  MoveL 647 to (-2817.75, 812.38, 1030.88) mm, rotated rx -103.17 ry -2.27 rz -179.99 deg; joints [-49.243, 2.601, 19.186, -115.031, 26.585, 9.042, -170]
  MoveL 648 to (-2817.75, 831.47, 992.27) mm, rotated rx -103.22 ry -3.45 rz -179.99 deg; joints [-48.787, 2.468, 20.52, -112.558, 24.893, 6.606, -170]
  MoveL 649 to (-2817.75, 844.77, 965.38) mm, rotated rx -103.26 ry -4.26 rz -179.99 deg; joints [-48.461, 2.4, 21.424, -110.645, 23.624, 4.8, -170]
  MoveL 650 to (-2817.75, 844.7, 935.74) mm, rotated rx -99.91 ry -3.73 rz -179.99 deg; joints [-48.443, 3.334, 22.932, -110.863, 27.836, -0.78, -170]
  MoveL 651 to (-2817.75, 844.62, 905.74) mm, rotated rx -96.49 ry -2.63 rz -179.99 deg; joints [-48.478, 4.555, 24.383, -112.634, 33.789, -5.769, -170]
  MoveL 652 to (-2817.75, 844.55, 875.74) mm, rotated rx -93.08 ry 1.03 rz 180 deg; joints [-48.572, 6.332, 25.892, -116.809, 44.188, -9.974, -170]
  MoveL 653 to (-2817.75, 844.47, 845.74) mm, rotated rx -89.7 ry 0.4 rz -179.6 deg; joints [-48.723, 7.85, 26.739, -119.615, 48.753, -14.494, -170]
  MoveL 654 to (-2817.75, 844.3, 816.11) mm, rotated rx -89.68 ry 0.41 rz -179.59 deg; joints [-48.729, 8.688, 27.11, -120.262, 50.179, -15.333, -170]
  MoveL 655 to (-2817.75, 844.12, 786.11) mm, rotated rx -89.67 ry 0.42 rz -179.58 deg; joints [-48.736, 9.565, 27.459, -120.936, 51.634, -16.183, -170]
  MoveL 656 to (-2817.75, 843.95, 756.11) mm, rotated rx -89.65 ry 0.43 rz -179.57 deg; joints [-48.743, 10.47, 27.78, -121.627, 53.1, -17.032, -170]
  MoveL 657 to (-2817.75, 843.77, 726.11) mm, rotated rx -89.64 ry 0.45 rz -179.56 deg; joints [-48.751, 11.401, 28.074, -122.336, 54.575, -17.882, -170]
  MoveL 658 to (-2817.75, 843.58, 696.48) mm, rotated rx -89.64 ry 0.45 rz -179.55 deg; joints [-48.758, 12.343, 28.335, -123.033, 56.012, -18.708, -170]
  MoveL 659 to (-2817.75, 843.38, 666.48) mm, rotated rx -89.64 ry 0.46 rz -179.54 deg; joints [-48.765, 13.323, 28.571, -123.754, 57.474, -19.544, -170]
  MoveL 660 to (-2817.75, 843.19, 636.48) mm, rotated rx -89.64 ry 0.47 rz -179.53 deg; joints [-48.773, 14.327, 28.78, -124.49, 58.942, -20.381, -170]
  MoveL 661 to (-2817.75, 843, 606.48) mm, rotated rx -89.64 ry 0.48 rz -179.52 deg; joints [-48.782, 15.356, 28.96, -125.239, 60.414, -21.219, -170]
  MoveL 662 to (-2817.75, 842.82, 569.69) mm, rotated rx -89.65 ry 0.48 rz -179.52 deg; joints [-48.789, 16.643, 29.145, -126.15, 62.194, -22.238, -170]
  MoveL 663 to (-2817.75, 842.68, 539.69) mm, rotated rx -89.66 ry 0.49 rz -179.51 deg; joints [-48.796, 17.718, 29.264, -126.907, 63.648, -23.068, -170]
  MoveL 664 to (-2817.75, 842.54, 509.69) mm, rotated rx -89.67 ry 0.49 rz -179.51 deg; joints [-48.803, 18.815, 29.354, -127.675, 65.102, -23.898, -170]
  MoveL 665 to (-2817.75, 842.4, 479.69) mm, rotated rx -89.68 ry 0.5 rz -179.5 deg; joints [-48.811, 19.933, 29.417, -128.453, 66.555, -24.728, -170]
  MoveL 666 to (-2817.75, 842.26, 449.69) mm, rotated rx -89.69 ry 0.5 rz -179.5 deg; joints [-48.819, 21.072, 29.451, -129.241, 68.007, -25.558, -170]
  MoveL 667 to (-2817.75, 842.12, 419.69) mm, rotated rx -89.7 ry 0.51 rz -179.5 deg; joints [-48.827, 22.229, 29.456, -130.038, 69.455, -26.387, -170]
  MoveL 668 to (-2817.75, 841.97, 389.69) mm, rotated rx -89.71 ry 0.51 rz -179.49 deg; joints [-48.836, 23.406, 29.433, -130.843, 70.899, -27.214, -170]
  MoveL 669 to (-2817.75, 841.83, 359.69) mm, rotated rx -89.73 ry 0.52 rz -179.49 deg; joints [-48.845, 24.599, 29.381, -131.655, 72.337, -28.04, -170]
  MoveL 670 to (-2817.75, 841.69, 329.69) mm, rotated rx -89.74 ry 0.52 rz -179.48 deg; joints [-48.855, 25.809, 29.301, -132.473, 73.767, -28.864, -170]
  MoveL 671 to (-2817.75, 841.54, 299.69) mm, rotated rx -89.75 ry 0.52 rz -179.48 deg; joints [-48.865, 27.035, 29.193, -133.296, 75.189, -29.685, -170]
  MoveL 672 to (-2817.75, 841.4, 269.7) mm, rotated rx -89.76 ry 0.53 rz -179.47 deg; joints [-48.876, 28.275, 29.056, -134.124, 76.601, -30.503, -170]
  MoveL 673 to (-2817.75, 841.26, 239.69) mm, rotated rx -89.75 ry -19.47 rz -179.55 deg; joints [-47.931, 25.571, 28.432, -109.218, 40.774, -38.612, -170]
  MoveL 674 to (-2817.75, 841.12, 209.69) mm, rotated rx -89.77 ry -19.46 rz -179.54 deg; joints [-47.933, 26.785, 28.338, -110.005, 42.222, -39.195, -170]
  MoveL 675 to (-2817.75, 841.08, 201.69) mm, rotated rx -89.77 ry -19.46 rz -179.54 deg; joints [-47.932, 27.113, 28.308, -110.208, 42.604, -39.356, -170]
  Set speed (1000.0 mm/s)
  MoveL 676 to (-2817.75, 841.08, 201.69) mm, rotated rx -89.77 ry -19.46 rz -179.54 deg; joints [-47.932, 27.113, 28.308, -110.208, 42.604, -39.356, -170]
  MoveL 677 to (-2818.68, 941.08, 201.3) mm, rotated rx -89.77 ry -19.46 rz -179.54 deg; joints [-46.038, 24.56, 32.438, -107.449, 43.1, -41.713, -170]
  Set speed (1000.0 mm/s)
  MoveL 678 to (-2898.69, 940.29, 202.16) mm, rotated rx -89.77 ry -19.46 rz -179.54 deg; joints [-49.032, 23.561, 34.225, -114.018, 46.527, -39.844, -170]
  MoveL 679 to (-2897.75, 840.3, 202.54) mm, rotated rx -89.77 ry -19.46 rz -179.54 deg; joints [-50.794, 26.176, 30.018, -116.607, 46.068, -37.565, -170]
  MoveL 680 to (-2897.75, 840.3, 202.54) mm, rotated rx -89.77 ry -19.46 rz -179.54 deg; joints [-50.794, 26.176, 30.018, -116.607, 46.068, -37.565, -170]
  Set speed (50.0 mm/s)
  MoveL 681 to (-2897.75, 840.33, 210.54) mm, rotated rx -89.77 ry -19.46 rz -179.54 deg; joints [-50.794, 25.842, 30.05, -116.45, 45.715, -37.364, -170]
  MoveL 682 to (-2897.75, 840.45, 240.54) mm, rotated rx -89.75 ry -19.46 rz -179.55 deg; joints [-50.792, 24.603, 30.15, -115.833, 44.378, -36.641, -170]
  MoveL 683 to (-2897.75, 840.57, 270.54) mm, rotated rx -89.74 ry -19.47 rz -179.56 deg; joints [-50.792, 23.378, 30.221, -115.24, 43.04, -35.89, -170]
  MoveL 684 to (-2897.75, 840.7, 300.54) mm, rotated rx -89.73 ry -19.47 rz -179.56 deg; joints [-50.792, 22.17, 30.264, -114.657, 41.697, -35.129, -170]
  MoveL 685 to (-2897.75, 840.81, 330.55) mm, rotated rx -89.74 ry 0.53 rz -179.48 deg; joints [-51.786, 24.874, 30.905, -137.578, 76.653, -28.084, -170]
  MoveL 686 to (-2897.75, 840.94, 360.54) mm, rotated rx -89.73 ry 0.52 rz -179.48 deg; joints [-51.777, 23.638, 30.987, -136.808, 75.263, -27.171, -170]
  MoveL 687 to (-2897.75, 841.02, 380.87) mm, rotated rx -89.72 ry 0.52 rz -179.48 deg; joints [-51.771, 22.81, 31.027, -136.292, 74.318, -26.55, -170]
  MoveL 688 to (-2897.75, 841.2, 410.87) mm, rotated rx -89.71 ry 0.52 rz -179.49 deg; joints [-51.761, 21.603, 31.063, -135.536, 72.922, -25.638, -170]
  MoveL 689 to (-2897.75, 841.38, 440.87) mm, rotated rx -89.7 ry 0.51 rz -179.49 deg; joints [-51.751, 20.414, 31.07, -134.791, 71.523, -24.724, -170]
  MoveL 690 to (-2897.75, 841.55, 470.87) mm, rotated rx -89.68 ry 0.51 rz -179.5 deg; joints [-51.742, 19.245, 31.049, -134.059, 70.124, -23.807, -170]
  MoveL 691 to (-2897.75, 841.73, 500.87) mm, rotated rx -89.67 ry 0.5 rz -179.5 deg; joints [-51.734, 18.096, 30.999, -133.341, 68.725, -22.888, -170]
  MoveL 692 to (-2897.75, 841.9, 530.87) mm, rotated rx -89.65 ry 0.5 rz -179.51 deg; joints [-51.726, 16.969, 30.92, -132.638, 67.328, -21.966, -170]
  MoveL 693 to (-2897.75, 842.07, 560.87) mm, rotated rx -89.64 ry 0.49 rz -179.51 deg; joints [-51.718, 15.864, 30.813, -131.95, 65.935, -21.042, -170]
  MoveL 694 to (-2897.75, 842.25, 590.87) mm, rotated rx -89.63 ry 0.48 rz -179.52 deg; joints [-51.711, 14.782, 30.677, -131.28, 64.547, -20.117, -170]
  MoveL 695 to (-2897.75, 842.37, 611.21) mm, rotated rx -89.62 ry 0.48 rz -179.52 deg; joints [-51.707, 14.062, 30.568, -130.835, 63.609, -19.488, -170]
  MoveL 696 to (-2897.75, 842.57, 641.21) mm, rotated rx -89.62 ry 0.47 rz -179.53 deg; joints [-51.699, 13.016, 30.385, -130.177, 62.209, -18.547, -170]
  MoveL 697 to (-2897.75, 842.78, 671.2) mm, rotated rx -89.62 ry 0.46 rz -179.54 deg; joints [-51.692, 11.994, 30.174, -129.54, 60.818, -17.604, -170]
  MoveL 698 to (-2897.75, 842.98, 701.2) mm, rotated rx -89.61 ry 0.46 rz -179.55 deg; joints [-51.685, 10.999, 29.935, -128.923, 59.438, -16.66, -170]
  MoveL 699 to (-2897.75, 843.19, 731.86) mm, rotated rx -89.61 ry 0.45 rz -179.55 deg; joints [-51.678, 10.01, 29.661, -128.315, 58.039, -15.693, -170]
  MoveL 700 to (-2897.75, 843.38, 761.86) mm, rotated rx -89.63 ry 0.44 rz -179.57 deg; joints [-51.671, 9.065, 29.363, -127.726, 56.658, -14.729, -170]
  MoveL 701 to (-2897.75, 843.57, 791.85) mm, rotated rx -89.64 ry 0.43 rz -179.58 deg; joints [-51.665, 8.149, 29.038, -127.162, 55.292, -13.763, -170]
  MoveL 702 to (-2897.75, 843.76, 821.85) mm, rotated rx -89.65 ry 0.41 rz -179.59 deg; joints [-51.659, 7.261, 28.685, -126.623, 53.941, -12.795, -170]
  MoveL 703 to (-2897.75, 843.96, 852.51) mm, rotated rx -89.67 ry 0.4 rz -179.6 deg; joints [-51.653, 6.383, 28.296, -126.1, 52.579, -11.802, -170]
  MoveL 704 to (-2897.75, 844.05, 882.51) mm, rotated rx -93.14 ry 0.91 rz 180 deg; joints [-51.496, 4.806, 27.427, -123.67, 48.036, -6.803, -170]
  MoveL 705 to (-2897.75, 844.14, 912.51) mm, rotated rx -96.65 ry -2.69 rz -179.99 deg; joints [-51.402, 3.012, 25.922, -121.089, 38.685, -1.519, -170]
  MoveL 706 to (-2897.75, 844.24, 942.51) mm, rotated rx -100.16 ry -3.78 rz -179.99 deg; joints [-51.372, 1.784, 24.461, -120.72, 33.653, 4.42, -170]
  MoveL 707 to (-2897.75, 844.33, 973.16) mm, rotated rx -103.72 ry -4.31 rz -179.99 deg; joints [-51.402, 0.829, 22.882, -121.934, 30.285, 11.118, -170]
  MoveL 708 to (-2897.75, 830.58, 999.82) mm, rotated rx -103.69 ry -3.5 rz -179.99 deg; joints [-51.725, 0.942, 21.926, -123.457, 31.388, 12.672, -170]
  MoveL 709 to (-2897.75, 809.97, 1039.78) mm, rotated rx -103.64 ry -2.29 rz -179.99 deg; joints [-52.194, 1.149, 20.461, -125.527, 32.941, 14.887, -170]
  MoveL 710 to (-2897.75, 796.37, 1066.52) mm, rotated rx -108.84 ry -1.41 rz -180 deg; joints [-52.753, 1.175, 17.955, -130.919, 33.223, 25.392, -170]
  MoveL 711 to (-2897.75, 775.99, 1106.6) mm, rotated rx -116.66 ry -0.72 rz -180 deg; joints [-53.755, 1.801, 13.687, -142.342, 36.014, 42.395, -170]
  MoveL 712 to (-2897.75, 762.7, 1133.49) mm, rotated rx -116.26 ry 0.34 rz 180 deg; joints [-54.078, 2.014, 12.796, -142.876, 37.16, 42.843, -170]
  MoveL 713 to (-2897.75, 749.89, 1159.4) mm, rotated rx -115.89 ry 1.39 rz 180 deg; joints [-54.38, 2.235, 11.926, -143.28, 38.216, 43.237, -170]
  MoveL 714 to (-2897.75, 746.94, 1165.63) mm, rotated rx -115.75 ry 1.69 rz 180 deg; joints [-54.45, 2.282, 11.747, -143.268, 38.475, 43.216, -170]
  Set speed (1000.0 mm/s)
  MoveL 715 to (-2897.75, 746.94, 1165.63) mm, rotated rx -115.75 ry 1.69 rz 180 deg; joints [-54.45, 2.282, 11.747, -143.268, 38.475, 43.216, -170]
  MoveL 716 to (-2899.02, 837.01, 1209.06) mm, rotated rx -115.75 ry 1.69 rz 180 deg; joints [-53.221, -1.859, 14.256, -141.506, 35.807, 44.207, -170]
  Set speed (1000.0 mm/s)
  MoveL 717 to (-2979.82, 828.97, 1222.94) mm, rotated rx -116.54 ry 2.68 rz 179.99 deg; joints [-56.639, -2.784, 14.766, -150.413, 43.399, 48.713, -170]
  MoveL 718 to (-2977.75, 739.51, 1178.3) mm, rotated rx -116.54 ry 2.68 rz 179.99 deg; joints [-57.642, 1.416, 12.276, -151.236, 45.388, 47.167, -170]
  MoveL 719 to (-2977.75, 739.51, 1178.3) mm, rotated rx -116.54 ry 2.68 rz 179.99 deg; joints [-57.642, 1.416, 12.276, -151.236, 45.388, 47.167, -170]
  Set speed (50.0 mm/s)
  MoveL 720 to (-2977.75, 743.33, 1170.64) mm, rotated rx -116.9 ry 1.76 rz 180 deg; joints [-57.513, 1.36, 12.335, -151.884, 44.805, 47.788, -170]
  MoveL 721 to (-2977.75, 757.4, 1143.51) mm, rotated rx -117.39 ry 0.32 rz 180 deg; joints [-57.172, 1.086, 13.2, -151.998, 43.61, 47.787, -170]
  MoveL 722 to (-2977.75, 771.22, 1116.88) mm, rotated rx -117.73 ry -0.71 rz -180 deg; joints [-56.858, 0.82, 14.158, -151.612, 42.569, 47.354, -170]
  MoveL 723 to (-2977.75, 779.23, 1101.8) mm, rotated rx -114.73 ry -0.91 rz -180 deg; joints [-56.469, 0.423, 15.935, -147.19, 41.112, 41.102, -170]
  MoveL 724 to (-2977.75, 793.31, 1075.31) mm, rotated rx -109.41 ry -1.43 rz -180 deg; joints [-55.836, -0.019, 18.855, -140.279, 39.466, 30.188, -170]
  MoveL 725 to (-2977.75, 807.39, 1048.82) mm, rotated rx -104.13 ry -2.31 rz -179.99 deg; joints [-55.283, -0.138, 21.477, -134.908, 38.92, 19.784, -170]
  MoveL 726 to (-2977.75, 815.48, 1033.78) mm, rotated rx -104.14 ry -2.76 rz -179.99 deg; joints [-55.114, -0.249, 22.065, -134.286, 38.393, 19.044, -170]
  MoveL 727 to (-2977.75, 829.69, 1007.36) mm, rotated rx -104.17 ry -3.56 rz -179.99 deg; joints [-54.811, -0.429, 23.083, -133.124, 37.432, 17.709, -170]
  MoveL 728 to (-2977.75, 843.89, 980.94) mm, rotated rx -104.2 ry -4.35 rz -179.99 deg; joints [-54.498, -0.589, 24.085, -131.869, 36.428, 16.329, -170]
  MoveL 729 to (-2977.75, 843.78, 949.27) mm, rotated rx -100.41 ry -3.82 rz -179.99 deg; joints [-54.457, 0.383, 25.761, -129.756, 39.228, 8.855, -170]
  MoveL 730 to (-2977.75, 843.66, 919.27) mm, rotated rx -96.8 ry -2.76 rz -179.99 deg; joints [-54.481, 1.615, 27.246, -129.178, 43.575, 2.269, -170]
  MoveL 731 to (-2977.75, 843.55, 889.27) mm, rotated rx -93.2 ry 0.78 rz 180 deg; joints [-54.569, 3.423, 28.761, -130.525, 52.047, -3.846, -170]
  MoveL 732 to (-2977.75, 843.44, 859.27) mm, rotated rx -89.64 ry 0.41 rz -179.6 deg; joints [-54.731, 5.056, 29.653, -132.597, 56.549, -9.299, -170]
  MoveL 733 to (-2977.75, 843.22, 827.6) mm, rotated rx -89.62 ry 0.42 rz -179.58 deg; joints [-54.735, 5.97, 30.06, -133.01, 57.842, -10.434, -170]
  MoveL 734 to (-2977.75, 843.02, 797.6) mm, rotated rx -89.61 ry 0.43 rz -179.57 deg; joints [-54.739, 6.868, 30.418, -133.433, 59.089, -11.505, -170]
  MoveL 735 to (-2977.75, 842.81, 767.6) mm, rotated rx -89.6 ry 0.44 rz -179.56 deg; joints [-54.744, 7.794, 30.748, -133.887, 60.356, -12.572, -170]
  MoveL 736 to (-2977.75, 842.61, 737.6) mm, rotated rx -89.59 ry 0.45 rz -179.55 deg; joints [-54.75, 8.75, 31.05, -134.37, 61.641, -13.636, -170]
  MoveL 737 to (-2977.75, 842.38, 705.93) mm, rotated rx -89.59 ry 0.46 rz -179.54 deg; joints [-54.756, 9.785, 31.337, -134.893, 62.992, -14.739, -170]
  MoveL 738 to (-2977.75, 842.16, 675.93) mm, rotated rx -89.59 ry 0.47 rz -179.53 deg; joints [-54.761, 10.794, 31.58, -135.416, 64.287, -15.781, -170]
  MoveL 739 to (-2977.75, 841.95, 645.94) mm, rotated rx -89.6 ry 0.48 rz -179.53 deg; joints [-54.768, 11.83, 31.795, -135.965, 65.597, -16.82, -170]
  MoveL 740 to (-2977.75, 841.73, 615.94) mm, rotated rx -89.6 ry 0.48 rz -179.52 deg; joints [-54.775, 12.893, 31.981, -136.537, 66.918, -17.856, -170]
  MoveL 741 to (-2977.75, 841.6, 593.66) mm, rotated rx -89.61 ry 0.49 rz -179.51 deg; joints [-54.779, 13.694, 32.101, -136.965, 67.89, -18.613, -170]
  MoveL 742 to (-2977.75, 841.41, 563.66) mm, rotated rx -89.62 ry 0.49 rz -179.51 deg; joints [-54.786, 14.794, 32.238, -137.56, 69.208, -19.63, -170]
  MoveL 743 to (-2977.75, 841.23, 533.66) mm, rotated rx -89.64 ry 0.5 rz -179.51 deg; joints [-54.792, 15.918, 32.346, -138.176, 70.533, -20.644, -170]
  MoveL 744 to (-2977.75, 841.05, 503.66) mm, rotated rx -89.65 ry 0.5 rz -179.5 deg; joints [-54.8, 17.065, 32.425, -138.812, 71.866, -21.655, -170]
  MoveL 745 to (-2977.75, 840.87, 473.66) mm, rotated rx -89.67 ry 0.51 rz -179.5 deg; joints [-54.808, 18.234, 32.475, -139.466, 73.203, -22.662, -170]
  MoveL 746 to (-2977.75, 840.68, 443.66) mm, rotated rx -89.68 ry 0.51 rz -179.49 deg; joints [-54.817, 19.425, 32.496, -140.138, 74.543, -23.665, -170]
  MoveL 747 to (-2977.75, 840.49, 413.67) mm, rotated rx -89.7 ry 0.52 rz -179.49 deg; joints [-54.826, 20.635, 32.488, -140.826, 75.886, -24.664, -170]
  MoveL 748 to (-2977.75, 840.31, 383.68) mm, rotated rx -89.71 ry 0.52 rz -179.48 deg; joints [-54.836, 21.864, 32.45, -141.528, 77.228, -25.659, -170]
  MoveL 749 to (-2977.75, 840.22, 361.39) mm, rotated rx -89.7 ry -19.48 rz -179.58 deg; joints [-53.805, 18.856, 31.81, -120.744, 43.029, -31.253, -170]
  MoveL 750 to (-2977.75, 840.1, 331.39) mm, rotated rx -89.71 ry -19.47 rz -179.57 deg; joints [-53.802, 20.05, 31.819, -121.094, 44.23, -32.192, -170]
  MoveL 751 to (-2977.75, 839.97, 301.39) mm, rotated rx -89.72 ry -19.47 rz -179.57 deg; joints [-53.8, 21.263, 31.798, -121.472, 45.44, -33.114, -170]
  MoveL 752 to (-2977.75, 839.84, 271.39) mm, rotated rx -89.73 ry -19.47 rz -179.56 deg; joints [-53.798, 22.495, 31.75, -121.875, 46.657, -34.019, -170]
  MoveL 753 to (-2977.75, 839.71, 241.39) mm, rotated rx -89.74 ry -19.46 rz -179.55 deg; joints [-53.797, 23.744, 31.672, -122.3, 47.878, -34.907, -170]
  MoveL 754 to (-2977.75, 839.58, 211.39) mm, rotated rx -89.75 ry -19.46 rz -179.55 deg; joints [-53.796, 25.01, 31.566, -122.744, 49.101, -35.779, -170]
  MoveL 755 to (-2977.75, 839.55, 203.39) mm, rotated rx -89.75 ry -19.46 rz -179.55 deg; joints [-53.795, 25.351, 31.533, -122.862, 49.427, -36.014, -170]
  Set speed (1000.0 mm/s)
  MoveL 756 to (-2977.75, 839.55, 203.39) mm, rotated rx -89.75 ry -19.46 rz -179.55 deg; joints [-53.795, 25.351, 31.533, -122.862, 49.427, -36.014, -170]
  MoveL 757 to (-2978.68, 939.54, 202.98) mm, rotated rx -89.75 ry -19.46 rz -179.55 deg; joints [-52.193, 22.678, 35.815, -120.489, 49.872, -38.211, -170]
  Set speed (1000.0 mm/s)
  MoveL 758 to (-3058.69, 938.8, 203.83) mm, rotated rx -89.75 ry -19.46 rz -179.54 deg; joints [-55.525, 21.905, 37.195, -126.964, 53.169, -36.713, -170]
  MoveL 759 to (-3057.75, 838.8, 204.24) mm, rotated rx -89.75 ry -19.46 rz -179.54 deg; joints [-56.937, 24.633, 32.844, -129.079, 52.722, -34.6, -170]
  MoveL 760 to (-3057.75, 838.8, 204.24) mm, rotated rx -89.75 ry -19.46 rz -179.54 deg; joints [-56.937, 24.633, 32.844, -129.079, 52.722, -34.6, -170]
  Set speed (50.0 mm/s)
  MoveL 761 to (-3057.75, 838.84, 212.24) mm, rotated rx -89.75 ry -19.46 rz -179.54 deg; joints [-56.939, 24.287, 32.878, -128.997, 52.425, -34.335, -170]
  MoveL 762 to (-3057.75, 838.97, 242.24) mm, rotated rx -89.73 ry -19.46 rz -179.56 deg; joints [-56.94, 23.001, 32.989, -128.679, 51.31, -33.367, -170]
  MoveL 763 to (-3057.75, 839.11, 272.24) mm, rotated rx -89.72 ry -19.46 rz -179.56 deg; joints [-56.943, 21.73, 33.072, -128.401, 50.204, -32.361, -170]
  MoveL 764 to (-3057.75, 839.24, 302.24) mm, rotated rx -89.71 ry -19.47 rz -179.57 deg; joints [-56.947, 20.477, 33.125, -128.153, 49.108, -31.335, -170]
  MoveL 765 to (-3057.75, 839.37, 332.24) mm, rotated rx -89.7 ry -19.47 rz -179.58 deg; joints [-56.952, 19.242, 33.149, -127.938, 48.026, -30.288, -170]
  MoveL 766 to (-3057.75, 839.5, 362.24) mm, rotated rx -89.69 ry -19.47 rz -179.58 deg; joints [-56.958, 18.028, 33.145, -127.758, 46.959, -29.22, -170]
  MoveL 767 to (-3057.75, 839.61, 386.45) mm, rotated rx -89.68 ry -19.48 rz -179.59 deg; joints [-56.963, 17.063, 33.12, -127.641, 46.112, -28.341, -170]
  MoveL 768 to (-3057.75, 839.8, 416.45) mm, rotated rx -89.67 ry -19.48 rz -179.6 deg; joints [-56.968, 15.888, 33.067, -127.521, 45.079, -27.245, -170]
  MoveL 769 to (-3057.75, 839.99, 446.45) mm, rotated rx -89.65 ry -19.49 rz -179.61 deg; joints [-56.974, 14.735, 32.985, -127.445, 44.069, -26.126, -170]
  MoveL 770 to (-3057.75, 840.17, 476.46) mm, rotated rx -89.65 ry 0.51 rz -179.49 deg; joints [-58.006, 17.35, 33.697, -144.988, 76.368, -21.607, -170]
  MoveL 771 to (-3057.75, 840.37, 506.45) mm, rotated rx -89.64 ry 0.5 rz -179.5 deg; joints [-57.998, 16.163, 33.647, -144.396, 75.101, -20.52, -170]
  MoveL 772 to (-3057.75, 840.56, 536.45) mm, rotated rx -89.62 ry 0.5 rz -179.5 deg; joints [-57.992, 14.999, 33.568, -143.824, 73.842, -19.428, -170]
  MoveL 773 to (-3057.75, 840.75, 566.45) mm, rotated rx -89.61 ry 0.49 rz -179.51 deg; joints [-57.986, 13.858, 33.459, -143.276, 72.591, -18.332, -170]
  MoveL 774 to (-3057.75, 840.94, 596.45) mm, rotated rx -89.59 ry 0.49 rz -179.51 deg; joints [-57.981, 12.742, 33.321, -142.75, 71.351, -17.232, -170]
  MoveL 775 to (-3057.75, 841.1, 620.66) mm, rotated rx -89.58 ry 0.49 rz -179.52 deg; joints [-57.977, 11.859, 33.189, -142.344, 70.359, -16.341, -170]
  MoveL 776 to (-3057.75, 841.32, 650.66) mm, rotated rx -89.58 ry 0.48 rz -179.52 deg; joints [-57.971, 10.784, 32.999, -141.85, 69.121, -15.221, -170]
  MoveL 777 to (-3057.75, 841.55, 680.66) mm, rotated rx -89.57 ry 0.47 rz -179.53 deg; joints [-57.966, 9.735, 32.782, -141.382, 67.898, -14.097, -170]
  MoveL 778 to (-3057.75, 841.78, 710.66) mm, rotated rx -89.57 ry 0.46 rz -179.54 deg; joints [-57.962, 8.715, 32.535, -140.943, 66.692, -12.969, -170]
  MoveL 779 to (-3057.75, 842.03, 743.35) mm, rotated rx -89.57 ry 0.45 rz -179.55 deg; joints [-57.958, 7.635, 32.234, -140.497, 65.398, -11.737, -170]
  MoveL 780 to (-3057.75, 842.24, 773.35) mm, rotated rx -89.58 ry 0.44 rz -179.56 deg; joints [-57.954, 6.671, 31.927, -140.106, 64.21, -10.587, -170]
  MoveL 781 to (-3057.75, 842.46, 803.35) mm, rotated rx -89.59 ry 0.43 rz -179.57 deg; joints [-57.95, 5.736, 31.592, -139.747, 63.043, -9.434, -170]
  MoveL 782 to (-3057.75, 842.68, 833.34) mm, rotated rx -89.6 ry 0.42 rz -179.58 deg; joints [-57.948, 4.832, 31.229, -139.42, 61.899, -8.276, -170]
  MoveL 783 to (-3057.75, 842.92, 866.03) mm, rotated rx -89.61 ry 0.41 rz -179.59 deg; joints [-57.946, 3.882, 30.803, -139.103, 60.68, -7.011, -170]
  MoveL 784 to (-3057.75, 843.05, 896.03) mm, rotated rx -93.26 ry 0.66 rz 180 deg; joints [-57.783, 2.196, 29.885, -137.36, 56.237, -1.135, -170]
  MoveL 785 to (-3057.75, 843.18, 926.03) mm, rotated rx -96.96 ry -2.82 rz -179.99 deg; joints [-57.701, 0.378, 28.352, -136.967, 48.516, 5.612, -170]
  MoveL 786 to (-3057.75, 843.31, 956.03) mm, rotated rx -100.67 ry -3.86 rz -179.99 deg; joints [-57.681, -0.854, 26.831, -138.196, 44.709, 12.647, -170]
  MoveL 787 to (-3057.75, 843.45, 988.71) mm, rotated rx -104.68 ry -4.39 rz -179.99 deg; joints [-57.73, -1.838, 25.045, -140.913, 42.337, 20.7, -170]
  MoveL 788 to (-3057.75, 828.79, 1014.88) mm, rotated rx -104.65 ry -3.61 rz -179.99 deg; joints [-58.024, -1.63, 23.999, -141.956, 43.271, 21.947, -170]
  MoveL 789 to (-3057.75, 814.12, 1041.05) mm, rotated rx -104.63 ry -2.83 rz -179.99 deg; joints [-58.31, -1.403, 22.938, -142.921, 44.165, 23.158, -170]
  MoveL 790 to (-3057.75, 804.62, 1058) mm, rotated rx -104.62 ry -2.32 rz -179.99 deg; joints [-58.49, -1.246, 22.243, -143.505, 44.723, 23.925, -170]
  MoveL 791 to (-3057.75, 790.06, 1084.22) mm, rotated rx -109.97 ry -1.45 rz -180 deg; joints [-59.019, -1.031, 19.507, -148.741, 45.467, 34.141, -170]
  MoveL 792 to (-3057.75, 775.49, 1110.45) mm, rotated rx -115.36 ry -0.93 rz -180 deg; joints [-59.617, -0.484, 16.462, -155.274, 47.204, 44.684, -170]
  MoveL 793 to (-3057.75, 766.07, 1127.43) mm, rotated rx -118.82 ry -0.69 rz -180 deg; joints [-60.03, 0.046, 14.35, -159.965, 48.881, 51.473, -170]
  MoveL 794 to (-3057.75, 751.73, 1153.78) mm, rotated rx -118.54 ry 0.3 rz 180 deg; joints [-60.331, 0.368, 13.325, -160.261, 49.85, 51.927, -170]
  MoveL 795 to (-3057.75, 736.24, 1182.24) mm, rotated rx -118.24 ry 1.4 rz 180 deg; joints [-60.647, 0.733, 12.204, -160.492, 50.847, 52.404, -170]
  MoveL 796 to (-3057.75, 731.39, 1191.44) mm, rotated rx -118.09 ry 1.82 rz 180 deg; joints [-60.748, 0.843, 11.877, -160.442, 51.17, 52.44, -170]
  Set speed (1000.0 mm/s)
  MoveL 797 to (-3057.75, 731.39, 1191.44) mm, rotated rx -118.09 ry 1.82 rz 180 deg; joints [-60.748, 0.843, 11.877, -160.442, 51.17, 52.44, -170]
  MoveL 798 to (-3059.23, 819.6, 1238.51) mm, rotated rx -118.09 ry 1.82 rz 180 deg; joints [-59.934, -3.333, 14.238, -160.411, 49.821, 54.432, -170]
  Set speed (1000.0 mm/s)
  MoveL 799 to (-3139.91, 809.88, 1253.7) mm, rotated rx -119.13 ry 2.56 rz 179.99 deg; joints [-63.457, -3.721, 13.98, -167.758, 56.791, 57.644, -170]
  MoveL 800 to (-3137.75, 722.53, 1205.08) mm, rotated rx -119.13 ry 2.56 rz 179.99 deg; joints [-64.034, 0.46, 11.689, -167.306, 57.626, 55.463, -170]
  MoveL 801 to (-3137.75, 722.53, 1205.08) mm, rotated rx -119.13 ry 2.56 rz 179.99 deg; joints [-64.034, 0.46, 11.689, -167.306, 57.626, 55.463, -170]
  Set speed (50.0 mm/s)
  MoveL 802 to (-3137.75, 728.58, 1194.21) mm, rotated rx -119.32 ry 1.88 rz 180 deg; joints [-63.898, 0.308, 12.054, -167.567, 57.175, 55.534, -170]
  MoveL 803 to (-3137.75, 745.65, 1164.3) mm, rotated rx -119.71 ry 0.28 rz 180 deg; joints [-63.531, -0.132, 13.179, -167.862, 55.968, 55.389, -170]
  MoveL 804 to (-3137.75, 760.52, 1138.25) mm, rotated rx -119.93 ry -0.68 rz -180 deg; joints [-63.248, -0.511, 14.272, -167.625, 55.053, 54.895, -170]
  MoveL 805 to (-3137.75, 771.56, 1119.21) mm, rotated rx -115.97 ry -0.95 rz -180 deg; joints [-62.826, -1.199, 16.758, -162.667, 53.137, 47.548, -170]
  MoveL 806 to (-3137.75, 786.61, 1093.26) mm, rotated rx -110.52 ry -1.47 rz -180 deg; joints [-62.281, -1.85, 19.918, -156.523, 51.338, 37.383, -170]
  MoveL 807 to (-3137.75, 801.66, 1067.31) mm, rotated rx -105.12 ry -2.34 rz -179.99 deg; joints [-61.792, -2.162, 22.76, -151.493, 50.446, 27.411, -170]
  MoveL 808 to (-3137.75, 812.76, 1048.3) mm, rotated rx -105.13 ry -2.9 rz -179.99 deg; joints [-61.606, -2.375, 23.577, -150.95, 49.855, 26.61, -170]
  MoveL 809 to (-3137.75, 827.89, 1022.4) mm, rotated rx -105.14 ry -3.67 rz -179.99 deg; joints [-61.345, -2.649, 24.679, -150.153, 49.018, 25.497, -170]
  MoveL 810 to (-3137.75, 843.01, 996.49) mm, rotated rx -105.16 ry -4.43 rz -179.99 deg; joints [-61.075, -2.906, 25.766, -149.289, 48.144, 24.359, -170]
  MoveL 811 to (-3137.75, 842.85, 962.79) mm, rotated rx -100.93 ry -3.9 rz -179.99 deg; joints [-61.026, -1.913, 27.672, -146.163, 50.171, 15.856, -170]
  MoveL 812 to (-3137.75, 842.7, 932.79) mm, rotated rx -97.12 ry -2.88 rz -179.99 deg; joints [-61.045, -0.684, 29.235, -144.491, 53.54, 8.514, -170]
  MoveL 813 to (-3137.75, 842.55, 902.79) mm, rotated rx -93.33 ry 0.55 rz 180 deg; joints [-61.122, 1.141, 30.794, -144.16, 60.612, 1.294, -170]
  MoveL 814 to (-3137.75, 842.4, 872.79) mm, rotated rx -89.57 ry 0.41 rz -179.59 deg; joints [-61.285, 2.875, 31.737, -145.608, 64.982, -4.966, -170]
  MoveL 815 to (-3137.75, 842.14, 839.09) mm, rotated rx -89.57 ry 0.42 rz -179.58 deg; joints [-61.284, 3.859, 32.184, -145.845, 66.123, -6.349, -170]
  MoveL 816 to (-3137.75, 841.91, 809.09) mm, rotated rx -89.56 ry 0.44 rz -179.57 deg; joints [-61.284, 4.768, 32.552, -146.092, 67.165, -7.576, -170]
  MoveL 817 to (-3137.75, 841.68, 779.09) mm, rotated rx -89.55 ry 0.45 rz -179.56 deg; joints [-61.285, 5.708, 32.892, -146.373, 68.232, -8.801, -170]
  MoveL 818 to (-3137.75, 841.44, 749.09) mm, rotated rx -89.54 ry 0.46 rz -179.55 deg; joints [-61.287, 6.679, 33.204, -146.686, 69.321, -10.023, -170]
  MoveL 819 to (-3137.75, 841.17, 715.39) mm, rotated rx -89.55 ry 0.47 rz -179.54 deg; joints [-61.289, 7.8, 33.519, -147.062, 70.548, -11.375, -170]
  MoveL 820 to (-3137.75, 840.94, 685.39) mm, rotated rx -89.55 ry 0.47 rz -179.53 deg; joints [-61.292, 8.83, 33.77, -147.429, 71.662, -12.575, -170]
  MoveL 821 to (-3137.75, 840.7, 655.39) mm, rotated rx -89.56 ry 0.48 rz -179.52 deg; joints [-61.295, 9.888, 33.991, -147.825, 72.794, -13.773, -170]
  MoveL 822 to (-3137.75, 840.46, 625.39) mm, rotated rx -89.56 ry 0.49 rz -179.51 deg; joints [-61.3, 10.974, 34.184, -148.25, 73.942, -14.967, -170]
  MoveL 823 to (-3137.75, 840.28, 599.24) mm, rotated rx -89.57 ry 0.49 rz -179.51 deg; joints [-61.302, 11.937, 34.329, -148.63, 74.939, -15.992, -170]
  MoveL 824 to (-3137.75, 840.08, 569.24) mm, rotated rx -89.59 ry 0.5 rz -179.51 deg; joints [-61.306, 13.066, 34.468, -149.091, 76.095, -17.165, -170]
  MoveL 825 to (-3137.75, 839.89, 539.24) mm, rotated rx -89.58 ry -19.5 rz -179.64 deg; joints [-60.303, 10.568, 33.688, -135.279, 45.87, -20.153, -170]
  MoveL 826 to (-3137.75, 839.7, 509.24) mm, rotated rx -89.6 ry -19.49 rz -179.63 deg; joints [-60.29, 11.659, 33.855, -135.047, 46.637, -21.452, -170]
  MoveL 827 to (-3137.75, 839.5, 479.24) mm, rotated rx -89.62 ry -19.49 rz -179.62 deg; joints [-60.277, 12.777, 33.993, -134.868, 47.441, -22.727, -170]
  MoveL 828 to (-3137.75, 839.3, 449.24) mm, rotated rx -89.64 ry -19.48 rz -179.61 deg; joints [-60.266, 13.92, 34.103, -134.74, 48.277, -23.978, -170]
  MoveL 829 to (-3137.75, 839.1, 419.24) mm, rotated rx -89.65 ry -19.48 rz -179.6 deg; joints [-60.256, 15.087, 34.185, -134.661, 49.144, -25.204, -170]
  MoveL 830 to (-3137.75, 838.9, 389.24) mm, rotated rx -89.67 ry -19.48 rz -179.59 deg; joints [-60.247, 16.278, 34.237, -134.627, 50.038, -26.408, -170]
  MoveL 831 to (-3137.75, 838.78, 363.08) mm, rotated rx -89.68 ry -19.47 rz -179.59 deg; joints [-60.238, 17.335, 34.262, -134.624, 50.837, -27.449, -170]
  MoveL 832 to (-3137.75, 838.64, 333.08) mm, rotated rx -89.69 ry -19.47 rz -179.58 deg; joints [-60.229, 18.567, 34.264, -134.661, 51.774, -28.621, -170]
  MoveL 833 to (-3137.75, 838.51, 303.08) mm, rotated rx -89.7 ry -19.47 rz -179.57 deg; joints [-60.221, 19.819, 34.236, -134.736, 52.732, -29.771, -170]
  MoveL 834 to (-3137.75, 838.37, 273.08) mm, rotated rx -89.71 ry -19.46 rz -179.57 deg; joints [-60.214, 21.091, 34.179, -134.849, 53.706, -30.898, -170]
  MoveL 835 to (-3137.75, 838.23, 243.08) mm, rotated rx -89.72 ry -19.46 rz -179.56 deg; joints [-60.208, 22.381, 34.094, -134.996, 54.696, -32.002, -170]
  MoveL 836 to (-3137.75, 838.09, 213.08) mm, rotated rx -89.73 ry -19.46 rz -179.55 deg; joints [-60.202, 23.687, 33.979, -135.174, 55.697, -33.085, -170]
  MoveL 837 to (-3137.75, 838.05, 204.08) mm, rotated rx -89.73 ry -19.46 rz -179.55 deg; joints [-60.2, 24.083, 33.939, -135.23, 55.999, -33.411, -170]
  Set speed (1000.0 mm/s)
  MoveL 838 to (-3137.75, 838.05, 204.08) mm, rotated rx -89.73 ry -19.46 rz -179.55 deg; joints [-60.2, 24.083, 33.939, -135.23, 55.999, -33.411, -170]
  MoveL 839 to (-3138.68, 938.05, 203.64) mm, rotated rx -89.73 ry -19.46 rz -179.55 deg; joints [-59.005, 21.312, 38.353, -133.416, 56.473, -35.446, -170]
  Set speed (1000.0 mm/s)
  MoveL 840 to (-3218.69, 937.3, 205.5) mm, rotated rx -89.73 ry -19.45 rz -179.55 deg; joints [-62.625, 20.748, 39.291, -139.871, 59.682, -34.217, -170]
  MoveL 841 to (-3217.75, 837.31, 205.93) mm, rotated rx -89.73 ry -19.45 rz -179.55 deg; joints [-63.575, 23.564, 34.823, -141.359, 59.177, -32.258, -170]
  MoveL 842 to (-3217.75, 837.31, 205.93) mm, rotated rx -89.73 ry -19.45 rz -179.55 deg; joints [-63.575, 23.564, 34.823, -141.359, 59.177, -32.258, -170]
  Set speed (50.0 mm/s)
  MoveL 843 to (-3217.75, 837.35, 213.93) mm, rotated rx -89.73 ry -19.45 rz -179.55 deg; joints [-63.578, 23.208, 34.859, -141.34, 58.939, -31.947, -170]
  MoveL 844 to (-3217.75, 837.49, 243.93) mm, rotated rx -89.71 ry -19.46 rz -179.56 deg; joints [-63.584, 21.889, 34.978, -141.263, 58.052, -30.802, -170]
  MoveL 845 to (-3217.75, 837.63, 273.93) mm, rotated rx -89.7 ry -19.46 rz -179.57 deg; joints [-63.594, 20.584, 35.066, -141.232, 57.181, -29.616, -170]
  MoveL 846 to (-3217.75, 837.77, 303.93) mm, rotated rx -89.69 ry -19.47 rz -179.57 deg; joints [-63.605, 19.298, 35.125, -141.238, 56.328, -28.408, -170]
  MoveL 847 to (-3217.75, 837.92, 333.93) mm, rotated rx -89.68 ry -19.47 rz -179.58 deg; joints [-63.617, 18.031, 35.155, -141.283, 55.495, -27.176, -170]
  MoveL 848 to (-3217.75, 838.06, 363.93) mm, rotated rx -89.67 ry -19.47 rz -179.59 deg; joints [-63.629, 16.785, 35.155, -141.368, 54.685, -25.922, -170]
  MoveL 849 to (-3217.75, 838.19, 392.03) mm, rotated rx -89.66 ry -19.47 rz -179.59 deg; joints [-63.642, 15.637, 35.129, -141.487, 53.95, -24.727, -170]
  MoveL 850 to (-3217.75, 838.4, 422.03) mm, rotated rx -89.64 ry -19.48 rz -179.6 deg; joints [-63.655, 14.434, 35.076, -141.647, 53.189, -23.442, -170]
  MoveL 851 to (-3217.75, 838.6, 452.03) mm, rotated rx -89.62 ry -19.48 rz -179.61 deg; joints [-63.67, 13.255, 34.994, -141.852, 52.458, -22.136, -170]
  MoveL 852 to (-3217.75, 838.81, 482.03) mm, rotated rx -89.6 ry -19.49 rz -179.63 deg; joints [-63.685, 12.101, 34.882, -142.105, 51.76, -20.807, -170]
  MoveL 853 to (-3217.75, 839.01, 512.03) mm, rotated rx -89.59 ry -19.49 rz -179.64 deg; joints [-63.702, 10.973, 34.742, -142.407, 51.095, -19.456, -170]
  MoveL 854 to (-3217.75, 839.22, 542.03) mm, rotated rx -89.57 ry -19.5 rz -179.65 deg; joints [-63.721, 9.872, 34.573, -142.76, 50.467, -18.084, -170]
  MoveL 855 to (-3217.75, 839.43, 572.03) mm, rotated rx -89.55 ry -19.5 rz -179.66 deg; joints [-63.741, 8.799, 34.376, -143.164, 49.877, -16.691, -170]
  MoveL 856 to (-3217.75, 839.63, 602.03) mm, rotated rx -89.53 ry -19.5 rz -179.67 deg; joints [-63.762, 7.754, 34.15, -143.621, 49.328, -15.277, -170]
  MoveL 857 to (-3217.75, 839.82, 630.12) mm, rotated rx -89.51 ry -19.51 rz -179.68 deg; joints [-63.783, 6.801, 33.912, -144.097, 48.852, -13.935, -170]
  MoveL 858 to (-3217.75, 840.06, 660.13) mm, rotated rx -89.54 ry 0.48 rz -179.52 deg; joints [-64.723, 9.154, 34.762, -153.876, 76.619, -12.5, -170]
  MoveL 859 to (-3217.75, 840.31, 690.12) mm, rotated rx -89.53 ry 0.48 rz -179.53 deg; joints [-64.721, 8.09, 34.537, -153.542, 75.582, -11.242, -170]
  MoveL 860 to (-3217.75, 840.57, 720.12) mm, rotated rx -89.53 ry 0.47 rz -179.53 deg; joints [-64.721, 7.054, 34.283, -153.237, 74.565, -9.982, -170]
  MoveL 861 to (-3217.75, 840.86, 754.84) mm, rotated rx -89.52 ry 0.46 rz -179.54 deg; joints [-64.721, 5.893, 33.953, -152.923, 73.413, -8.52, -170]
  MoveL 862 to (-3217.75, 841.1, 784.84) mm, rotated rx -89.53 ry 0.45 rz -179.55 deg; joints [-64.721, 4.919, 33.636, -152.673, 72.423, -7.241, -170]
  MoveL 863 to (-3217.75, 841.35, 814.84) mm, rotated rx -89.53 ry 0.44 rz -179.56 deg; joints [-64.722, 3.975, 33.29, -152.456, 71.456, -5.96, -170]
  MoveL 864 to (-3217.75, 841.6, 844.84) mm, rotated rx -89.54 ry 0.43 rz -179.57 deg; joints [-64.724, 3.064, 32.917, -152.271, 70.514, -4.678, -170]
  MoveL 865 to (-3217.75, 841.88, 879.55) mm, rotated rx -89.54 ry 0.42 rz -179.59 deg; joints [-64.727, 2.049, 32.45, -152.098, 69.456, -3.192, -170]
  MoveL 866 to (-3217.75, 842.05, 909.55) mm, rotated rx -93.39 ry 0.44 rz 180 deg; joints [-64.566, 0.272, 31.481, -150.904, 65.169, 3.41, -170]
  MoveL 867 to (-3217.75, 842.22, 939.55) mm, rotated rx -97.28 ry -2.94 rz -179.99 deg; joints [-64.493, -1.557, 29.891, -151.769, 58.658, 10.972, -170]
  MoveL 868 to (-3217.75, 842.38, 969.55) mm, rotated rx -101.18 ry -3.94 rz -179.99 deg; joints [-64.471, -2.782, 28.284, -153.731, 55.653, 18.519, -170]
  MoveL 869 to (-3217.75, 842.57, 1004.27) mm, rotated rx -105.65 ry -4.47 rz -179.99 deg; joints [-64.511, -3.779, 26.252, -157.129, 53.912, 27.379, -170]
  MoveL 870 to (-3217.75, 826.98, 1029.9) mm, rotated rx -105.64 ry -3.72 rz -179.99 deg; joints [-64.75, -3.474, 25.126, -157.837, 54.73, 28.431, -170]
  MoveL 871 to (-3217.75, 811.39, 1055.53) mm, rotated rx -105.63 ry -2.97 rz -179.99 deg; joints [-64.98, -3.153, 23.986, -158.485, 55.513, 29.464, -170]
  MoveL 872 to (-3217.75, 798.48, 1076.76) mm, rotated rx -105.62 ry -2.35 rz -179.99 deg; joints [-65.165, -2.874, 23.033, -158.98, 56.135, 30.307, -170]
  MoveL 873 to (-3217.75, 782.95, 1102.42) mm, rotated rx -111.07 ry -1.49 rz -180 deg; joints [-65.599, -2.466, 20.092, -163.761, 57.135, 40.003, -170]
  MoveL 874 to (-3217.75, 767.41, 1128.08) mm, rotated rx -116.55 ry -0.97 rz -180 deg; joints [-66.076, -1.716, 16.83, -169.519, 58.969, 49.793, -170]
  MoveL 875 to (-3217.75, 754.54, 1149.34) mm, rotated rx -121.06 ry -0.67 rz -180 deg; joints [-66.489, -0.845, 13.93, -174.739, 61.138, 57.717, -170]
  MoveL 876 to (-3217.75, 739.14, 1175.08) mm, rotated rx -120.89 ry 0.25 rz 180 deg; joints [-66.749, -0.408, 12.769, -174.936, 62.008, 58.259, -170]
  MoveL 877 to (-3217.75, 720.31, 1206.54) mm, rotated rx -120.7 ry 1.39 rz 180 deg; joints [-67.055, 0.146, 11.332, -175.102, 63.015, 58.925, -170]
  MoveL 878 to (-3217.75, 712.89, 1219.19) mm, rotated rx -120.57 ry 1.93 rz 180 deg; joints [-67.181, 0.363, 10.788, -175.046, 63.419, 59.099, -170]
  Set speed (1000.0 mm/s)
  MoveL 879 to (-3217.75, 712.89, 1219.19) mm, rotated rx -120.57 ry 1.93 rz 180 deg; joints [-67.181, 0.363, 10.788, -175.046, 63.419, 59.099, -170]
  MoveL 880 to (-3219.45, 798.99, 1270.03) mm, rotated rx -120.57 ry 1.93 rz 180 deg; joints [-66.793, -3.761, 12.942, -175.911, 63.089, 61.403, -170]
  Set speed (1000.0 mm/s)
  MoveL 881 to (-3299.96, 787.41, 1286.41) mm, rotated rx -121.79 ry 2.42 rz 179.99 deg; joints [-70.276, -3.576, 11.955, -182.436, 69.768, 63.717, -170]
  MoveL 882 to (-3297.75, 702.41, 1233.78) mm, rotated rx -121.79 ry 2.42 rz 179.99 deg; joints [-70.441, 0.497, 9.906, -181.294, 69.652, 61.416, -170]
  MoveL 883 to (-3297.75, 702.41, 1233.78) mm, rotated rx -121.79 ry 2.42 rz 179.99 deg; joints [-70.441, 0.497, 9.906, -181.294, 69.652, 61.416, -170]
  Set speed (50.0 mm/s)
  MoveL 884 to (-3297.75, 711.41, 1219.24) mm, rotated rx -121.86 ry 1.98 rz 180 deg; joints [-70.331, 0.206, 10.625, -181.226, 69.273, 61.058, -170]
  MoveL 885 to (-3297.75, 732.18, 1186.12) mm, rotated rx -122.09 ry 0.23 rz 180 deg; joints [-69.961, -0.456, 12.101, -181.58, 67.992, 60.609, -170]
  MoveL 886 to (-3297.75, 748.11, 1160.7) mm, rotated rx -122.2 ry -0.66 rz -180 deg; joints [-69.73, -0.951, 13.328, -181.413, 67.162, 60.012, -170]
  MoveL 887 to (-3297.75, 761.95, 1138.82) mm, rotated rx -119.85 ry -0.98 rz -180 deg; joints [-69.481, -1.692, 15.482, -178.569, 65.691, 55.7, -170]
  MoveL 888 to (-3297.75, 777.99, 1113.46) mm, rotated rx -117.11 ry -1.41 rz -180 deg; joints [-69.188, -2.456, 17.897, -175.367, 64.161, 50.594, -170]
  MoveL 889 to (-3297.75, 794.02, 1088.11) mm, rotated rx -114.35 ry -1.93 rz -180 deg; joints [-68.893, -3.114, 20.215, -172.313, 62.823, 45.407, -170]
  MoveL 890 to (-3297.75, 810.06, 1062.76) mm, rotated rx -111.6 ry -2.59 rz -179.99 deg; joints [-68.598, -3.663, 22.429, -169.458, 61.663, 40.183, -170]
  MoveL 891 to (-3297.75, 826.1, 1037.4) mm, rotated rx -108.86 ry -3.42 rz -179.99 deg; joints [-68.305, -4.105, 24.53, -166.847, 60.64, 34.969, -170]
  MoveL 892 to (-3297.75, 842.13, 1012.05) mm, rotated rx -106.14 ry -4.51 rz -179.99 deg; joints [-68.013, -4.447, 26.505, -164.521, 59.671, 29.815, -170]
  MoveL 893 to (-3297.75, 841.92, 976.31) mm, rotated rx -101.43 ry -3.97 rz -179.99 deg; joints [-67.99, -3.449, 28.668, -160.952, 61.17, 20.662, -170]
  MoveL 894 to (-3297.75, 841.73, 946.31) mm, rotated rx -97.43 ry -2.99 rz -179.99 deg; joints [-68.021, -2.23, 30.32, -158.816, 63.871, 12.988, -170]
  MoveL 895 to (-3297.75, 841.55, 916.31) mm, rotated rx -93.45 ry 0.34 rz 180 deg; joints [-68.094, -0.401, 31.942, -157.573, 69.899, 5.188, -170]
  MoveL 896 to (-3297.75, 841.36, 886.32) mm, rotated rx -89.51 ry 0.42 rz -179.58 deg; joints [-68.252, 1.416, 32.936, -158.56, 74.097, -1.713, -170]
  MoveL 897 to (-3297.75, 841.05, 850.58) mm, rotated rx -89.51 ry 0.43 rz -179.57 deg; joints [-68.246, 2.459, 33.424, -158.683, 75.069, -3.288, -170]
  MoveL 898 to (-3297.75, 840.78, 820.59) mm, rotated rx -89.5 ry 0.44 rz -179.56 deg; joints [-68.242, 3.37, 33.802, -158.821, 75.912, -4.61, -170]
  MoveL 899 to (-3297.75, 840.52, 790.6) mm, rotated rx -89.5 ry 0.45 rz -179.55 deg; joints [-68.239, 4.314, 34.152, -158.989, 76.779, -5.933, -170]
  MoveL 900 to (-3297.75, 840.27, 760.58) mm, rotated rx -89.47 ry -19.54 rz -179.72 deg; joints [-67.427, 2.229, 33.144, -154.537, 52.573, -5.683, -170]
  MoveL 901 to (-3297.75, 839.96, 724.85) mm, rotated rx -89.47 ry -19.53 rz -179.71 deg; joints [-67.389, 3.299, 33.589, -153.619, 52.835, -7.508, -170]
  MoveL 902 to (-3297.75, 839.7, 694.85) mm, rotated rx -89.48 ry -19.52 rz -179.7 deg; joints [-67.359, 4.232, 33.932, -152.898, 53.103, -9.029, -170]
  MoveL 903 to (-3297.75, 839.44, 664.85) mm, rotated rx -89.49 ry -19.51 rz -179.69 deg; joints [-67.331, 5.197, 34.247, -152.224, 53.414, -10.538, -170]
  MoveL 904 to (-3297.75, 839.18, 634.85) mm, rotated rx -89.5 ry -19.51 rz -179.68 deg; joints [-67.304, 6.193, 34.533, -151.597, 53.767, -12.034, -170]
  MoveL 905 to (-3297.75, 838.97, 604.81) mm, rotated rx -89.51 ry -19.5 rz -179.67 deg; joints [-67.277, 7.216, 34.792, -151.014, 54.149, -13.501, -170]
  MoveL 906 to (-3297.75, 838.76, 574.82) mm, rotated rx -89.53 ry -19.5 rz -179.66 deg; joints [-67.251, 8.266, 35.022, -150.478, 54.571, -14.952, -170]
  MoveL 907 to (-3297.75, 838.55, 544.82) mm, rotated rx -89.55 ry -19.49 rz -179.65 deg; joints [-67.227, 9.346, 35.223, -149.99, 55.032, -16.386, -170]
  MoveL 908 to (-3297.75, 838.33, 514.82) mm, rotated rx -89.57 ry -19.49 rz -179.64 deg; joints [-67.204, 10.454, 35.395, -149.547, 55.529, -17.804, -170]
  MoveL 909 to (-3297.75, 838.12, 484.82) mm, rotated rx -89.59 ry -19.49 rz -179.63 deg; joints [-67.183, 11.589, 35.538, -149.151, 56.063, -19.204, -170]
  MoveL 910 to (-3297.75, 837.91, 454.82) mm, rotated rx -89.61 ry -19.48 rz -179.62 deg; joints [-67.163, 12.75, 35.651, -148.8, 56.63, -20.586, -170]
  MoveL 911 to (-3297.75, 837.69, 424.82) mm, rotated rx -89.63 ry -19.48 rz -179.61 deg; joints [-67.144, 13.937, 35.735, -148.493, 57.23, -21.948, -170]
  MoveL 912 to (-3297.75, 837.48, 394.82) mm, rotated rx -89.65 ry -19.47 rz -179.6 deg; joints [-67.127, 15.148, 35.79, -148.23, 57.86, -23.291, -170]
  MoveL 913 to (-3297.75, 837.33, 364.78) mm, rotated rx -89.66 ry -19.47 rz -179.59 deg; joints [-67.109, 16.384, 35.818, -148, 58.517, -24.629, -170]
  MoveL 914 to (-3297.75, 837.19, 334.78) mm, rotated rx -89.67 ry -19.47 rz -179.58 deg; joints [-67.093, 17.641, 35.817, -147.811, 59.2, -25.943, -170]
  MoveL 915 to (-3297.75, 837.04, 304.78) mm, rotated rx -89.68 ry -19.46 rz -179.58 deg; joints [-67.077, 18.918, 35.786, -147.663, 59.908, -27.237, -170]
  MoveL 916 to (-3297.75, 836.89, 274.78) mm, rotated rx -89.69 ry -19.46 rz -179.57 deg; joints [-67.063, 20.215, 35.726, -147.553, 60.638, -28.508, -170]
  MoveL 917 to (-3297.75, 836.75, 244.78) mm, rotated rx -89.7 ry -19.46 rz -179.56 deg; joints [-67.05, 21.531, 35.636, -147.48, 61.387, -29.757, -170]
  MoveL 918 to (-3297.75, 836.6, 214.78) mm, rotated rx -89.72 ry -19.46 rz -179.56 deg; joints [-67.037, 22.865, 35.516, -147.442, 62.154, -30.982, -170]
  MoveL 919 to (-3297.75, 836.56, 206.78) mm, rotated rx -89.72 ry -19.46 rz -179.56 deg; joints [-67.034, 23.224, 35.479, -147.435, 62.361, -31.31, -170]
  Set speed (1000.0 mm/s)
  MoveL 920 to (-3297.75, 836.56, 206.78) mm, rotated rx -89.72 ry -19.46 rz -179.56 deg; joints [-67.034, 23.224, 35.479, -147.435, 62.361, -31.31, -170]
  MoveL 921 to (-3298.68, 936.56, 206.31) mm, rotated rx -89.72 ry -19.46 rz -179.56 deg; joints [-66.351, 20.379, 39.988, -146.303, 62.921, -33.208, -170]
  Set speed (1000.0 mm/s)
  MoveL 922 to (-3378.66, 936.76, 380.81) mm, rotated rx -89.66 ry -19.47 rz -179.59 deg; joints [-70.266, 12.017, 40.791, -153.729, 62.12, -24.131, -170]
  MoveL 923 to (-3377.75, 836.76, 381.38) mm, rotated rx -89.66 ry -19.47 rz -179.59 deg; joints [-70.665, 15.478, 36.237, -154.686, 62.05, -22.819, -170]
  MoveL 924 to (-3377.75, 836.76, 381.38) mm, rotated rx -89.66 ry -19.47 rz -179.59 deg; joints [-70.665, 15.478, 36.237, -154.686, 62.05, -22.819, -170]
  Set speed (50.0 mm/s)
  MoveL 925 to (-3377.75, 836.82, 389.38) mm, rotated rx -89.66 ry -19.47 rz -179.59 deg; joints [-70.671, 15.147, 36.229, -154.775, 61.911, -22.447, -170]
  MoveL 926 to (-3377.75, 837.04, 419.38) mm, rotated rx -89.62 ry -19.48 rz -179.61 deg; joints [-70.689, 13.928, 36.182, -155.088, 61.393, -21.097, -170]
  MoveL 927 to (-3377.75, 837.26, 449.38) mm, rotated rx -89.6 ry -19.48 rz -179.62 deg; joints [-70.711, 12.73, 36.104, -155.464, 60.911, -19.702, -170]
  MoveL 928 to (-3377.75, 837.48, 479.37) mm, rotated rx -89.59 ry -19.49 rz -179.63 deg; joints [-70.734, 11.557, 35.995, -155.88, 60.46, -18.291, -170]
  MoveL 929 to (-3377.75, 837.7, 509.37) mm, rotated rx -89.57 ry -19.49 rz -179.64 deg; joints [-70.759, 10.41, 35.857, -156.337, 60.042, -16.865, -170]
  MoveL 930 to (-3377.75, 837.92, 539.37) mm, rotated rx -89.55 ry -19.49 rz -179.65 deg; joints [-70.785, 9.291, 35.69, -156.835, 59.657, -15.425, -170]
  MoveL 931 to (-3377.75, 838.14, 569.37) mm, rotated rx -89.53 ry -19.5 rz -179.66 deg; joints [-70.812, 8.2, 35.492, -157.373, 59.308, -13.972, -170]
  MoveL 932 to (-3377.75, 838.36, 599.37) mm, rotated rx -89.52 ry -19.5 rz -179.67 deg; joints [-70.841, 7.138, 35.266, -157.952, 58.994, -12.507, -170]
  MoveL 933 to (-3377.75, 838.58, 629.37) mm, rotated rx -89.5 ry -19.51 rz -179.68 deg; joints [-70.871, 6.106, 35.011, -158.571, 58.717, -11.032, -170]
  MoveL 934 to (-3377.75, 838.8, 659.37) mm, rotated rx -89.48 ry -19.51 rz -179.69 deg; joints [-70.902, 5.105, 34.727, -159.229, 58.478, -9.548, -170]
  MoveL 935 to (-3377.75, 839.02, 689.37) mm, rotated rx -89.46 ry -19.52 rz -179.7 deg; joints [-70.935, 4.134, 34.414, -159.925, 58.276, -8.056, -170]
  MoveL 936 to (-3377.75, 839.22, 716.03) mm, rotated rx -89.45 ry -19.52 rz -179.71 deg; joints [-70.965, 3.298, 34.112, -160.576, 58.129, -6.725, -170]
  MoveL 937 to (-3377.75, 839.49, 746.03) mm, rotated rx -89.45 ry -19.53 rz -179.72 deg; joints [-70.998, 2.381, 33.746, -161.345, 57.985, -5.194, -170]
  MoveL 938 to (-3377.75, 839.77, 776.03) mm, rotated rx -89.45 ry -19.54 rz -179.73 deg; joints [-71.033, 1.496, 33.351, -162.151, 57.88, -3.659, -170]
  MoveL 939 to (-3377.75, 840.14, 817.3) mm, rotated rx -89.45 ry -19.55 rz -179.74 deg; joints [-71.083, 0.332, 32.762, -163.317, 57.801, -1.543, -170]
  MoveL 940 to (-3377.75, 840.42, 847.29) mm, rotated rx -89.46 ry -19.56 rz -179.75 deg; joints [-71.119, -0.476, 32.301, -164.202, 57.782, 0.006, -170]
  MoveL 941 to (-3377.75, 840.69, 877.29) mm, rotated rx -89.47 ry -19.57 rz -179.76 deg; joints [-71.156, -1.251, 31.812, -165.12, 57.801, 1.555, -170]
  MoveL 942 to (-3377.75, 841.07, 918.56) mm, rotated rx -89.48 ry -19.59 rz -179.77 deg; joints [-71.209, -2.263, 31.095, -166.431, 57.891, 3.683, -170]
  MoveL 943 to (-3377.75, 841.25, 948.56) mm, rotated rx -94.55 ry -1.26 rz -180 deg; joints [-71.669, -1.891, 31.411, -164.608, 72.303, 9.529, -170]
  MoveL 944 to (-3377.75, 841.44, 978.56) mm, rotated rx -99.66 ry -3.65 rz -179.99 deg; joints [-71.583, -3.577, 29.472, -166.857, 67.635, 18.972, -170]
  MoveL 945 to (-3377.75, 841.69, 1019.83) mm, rotated rx -106.64 ry -4.54 rz -179.99 deg; joints [-71.555, -4.903, 26.53, -171.532, 65.431, 31.712, -170]
  MoveL 946 to (-3377.75, 825.19, 1044.88) mm, rotated rx -109.35 ry -3.47 rz -179.99 deg; joints [-71.787, -4.496, 24.501, -173.658, 66.388, 36.699, -170]
  MoveL 947 to (-3377.75, 808.68, 1069.93) mm, rotated rx -112.1 ry -2.65 rz -179.99 deg; joints [-72.018, -3.99, 22.349, -176.048, 67.398, 41.731, -170]
  MoveL 948 to (-3377.75, 792.18, 1094.98) mm, rotated rx -114.86 ry -2 rz -180 deg; joints [-72.249, -3.378, 20.084, -178.667, 68.536, 46.76, -170]
  MoveL 949 to (-3377.75, 775.67, 1120.03) mm, rotated rx -117.63 ry -1.48 rz -180 deg; joints [-72.479, -2.659, 17.715, -181.47, 69.839, 51.743, -170]
  MoveL 950 to (-3377.75, 759.16, 1145.08) mm, rotated rx -120.38 ry -1.04 rz -180 deg; joints [-72.705, -1.836, 15.251, -184.415, 71.322, 56.644, -170]
  MoveL 951 to (-3377.74, 741.21, 1172.34) mm, rotated rx -123.35 ry -0.65 rz -180 deg; joints [-72.946, -0.827, 12.473, -187.728, 73.136, 61.842, -170]
  MoveL 952 to (-3377.74, 724.79, 1197.44) mm, rotated rx -123.27 ry 0.26 rz 180 deg; joints [-73.152, -0.28, 11.199, -187.815, 73.95, 62.449, -170]
  MoveL 953 to (-3377.74, 708.37, 1222.55) mm, rotated rx -123.19 ry 1.16 rz 180 deg; joints [-73.351, 0.281, 9.911, -187.859, 74.725, 63.067, -170]
  MoveL 954 to (-3377.74, 691.95, 1247.66) mm, rotated rx -123.13 ry 2.08 rz 180 deg; joints [-73.541, 0.854, 8.607, -187.861, 75.46, 63.698, -170]
  MoveL 955 to (-3377.74, 691.13, 1248.91) mm, rotated rx -123.12 ry 2.12 rz 180 deg; joints [-73.551, 0.883, 8.542, -187.86, 75.495, 63.73, -170]
  Set speed (1000.0 mm/s)
  MoveL 956 to (-3377.74, 691.13, 1248.91) mm, rotated rx -123.12 ry 2.12 rz 180 deg; joints [-73.551, 0.883, 8.542, -187.86, 75.495, 63.73, -170]
  MoveL 957 to (-3379.76, 774.87, 1303.51) mm, rotated rx -125.21 ry 18.73 rz 168.61 deg; joints [-71.519, -5.043, 15.187, -153.347, 58.212, 60.569, -170]
  Set speed (1000.0 mm/s)
  MoveL 958 to (-3460.49, 761.22, 1320.93) mm, rotated rx -126.73 ry 19.11 rz 168.18 deg; joints [-75.048, -4.482, 13.841, -160.128, 63.919, 64.662, -170]
  MoveL 959 to (-3457.75, 678.76, 1264.42) mm, rotated rx -126.73 ry 19.11 rz 168.18 deg; joints [-74.94, -0.426, 12.001, -159.282, 64.48, 62.162, -170]
  MoveL 960 to (-3457.75, 678.76, 1264.42) mm, rotated rx -126.73 ry 19.11 rz 168.18 deg; joints [-74.94, -0.426, 12.001, -159.282, 64.48, 62.162, -170]
  Set speed (50.0 mm/s)
  MoveL 961 to (-3457.75, 682.86, 1258.44) mm, rotated rx -126.59 ry 18.48 rz 168.22 deg; joints [-74.861, -0.585, 12.261, -159.539, 64.152, 61.976, -170]
  MoveL 962 to (-3457.75, 699.84, 1233.71) mm, rotated rx -126.38 ry 17.43 rz 168.29 deg; joints [-74.706, -1.175, 13.561, -159.739, 63.736, 61.066, -170]
  MoveL 963 to (-3457.75, 716.82, 1208.98) mm, rotated rx -126.21 ry 16.59 rz 168.34 deg; joints [-74.569, -1.745, 14.876, -159.792, 63.405, 60.138, -170]
  MoveL 964 to (-3457.75, 722.48, 1200.73) mm, rotated rx -126.15 ry 16.31 rz 168.36 deg; joints [-74.522, -1.932, 15.31, -159.801, 63.285, 59.83, -170]
  MoveL 965 to (-3457.75, 733.8, 1184.24) mm, rotated rx -126.05 ry 15.74 rz 168.39 deg; joints [-74.425, -2.303, 16.175, -159.804, 63.032, 59.214, -170]
  MoveL 966 to (-3457.75, 742.26, 1171.91) mm, rotated rx -124.63 ry 15.85 rz 168.79 deg; joints [-74.365, -2.664, 17.377, -159.108, 63.553, 56.721, -170]
  MoveL 967 to (-3457.75, 756.4, 1151.3) mm, rotated rx -122.25 ry 15.97 rz 169.49 deg; joints [-74.272, -3.205, 19.334, -158.165, 64.598, 52.589, -170]
  MoveL 968 to (-3457.75, 773.37, 1126.56) mm, rotated rx -125.82 ry 15.21 rz 168.45 deg; joints [-74.26, -3.496, 19.397, -159.117, 63.17, 56.714, -170]
  MoveL 969 to (-3457.75, 779.03, 1118.31) mm, rotated rx -125.8 ry 15.13 rz 168.46 deg; joints [-74.236, -3.658, 19.845, -159.023, 63.187, 56.381, -170]
  MoveL 970 to (-3457.75, 790.34, 1101.82) mm, rotated rx -125.78 ry 14.99 rz 168.47 deg; joints [-74.189, -3.978, 20.737, -158.834, 63.226, 55.713, -170]
  MoveL 971 to (-3457.75, 807.31, 1077.09) mm, rotated rx -129.68 ry 27.82 rz 167.08 deg; joints [-75.817, -3.423, 23.465, -155.667, 74.263, 55.525, -170]
  MoveL 972 to (-3457.75, 812.97, 1068.84) mm, rotated rx -140.04 ry 42.54 rz 149.69 deg; joints [-72.268, -4.845, 26.863, -122.733, 63.089, 49.899, -170]
  MoveL 973 to (-3457.75, 824.28, 1052.34) mm, rotated rx -140.82 ry 43.24 rz 149.18 deg; joints [-72.308, -5.004, 27.765, -123.024, 64.435, 49.883, -170]
  MoveL 974 to (-3457.75, 841.26, 1027.61) mm, rotated rx -89.39 ry -21.16 rz 178.64 deg; joints [-74.151, -5.171, 29.25, -173.097, 59.461, 9.671, -170]
  MoveL 975 to (-3457.75, 841.03, 997.35) mm, rotated rx -89.39 ry -20.97 rz 178.82 deg; joints [-74.2, -4.515, 29.873, -172.395, 59.724, 8.138, -170]
  MoveL 976 to (-3457.75, 840.85, 972.35) mm, rotated rx -89.39 ry -20.61 rz 179.18 deg; joints [-74.355, -3.882, 30.349, -172.35, 60.64, 6.867, -170]
  MoveL 977 to (-3457.75, 840.66, 947.35) mm, rotated rx -89.4 ry -19.52 rz -179.73 deg; joints [-74.903, -2.985, 30.731, -174.126, 63.922, 5.575, -170]
  MoveL 978 to (-3457.75, 840.48, 922.35) mm, rotated rx -92.95 ry -18.14 rz -178.99 deg; joints [-74.9, -2.761, 30.567, -175.513, 64.885, 9.495, -170]
  MoveL 979 to (-3457.75, 840.3, 897.35) mm, rotated rx -89.42 ry -19.57 rz -179.77 deg; joints [-74.802, -1.833, 31.643, -172.456, 63.459, 3.146, -170]
  MoveL 980 to (-3457.75, 840.14, 881.57) mm, rotated rx -89.42 ry -19.57 rz -179.77 deg; joints [-74.782, -1.441, 31.913, -171.983, 63.394, 2.363, -170]
  MoveL 981 to (-3457.75, 839.9, 856.57) mm, rotated rx -89.42 ry -19.56 rz -179.76 deg; joints [-74.749, -0.801, 32.327, -171.245, 63.308, 1.12, -170]
  MoveL 982 to (-3457.75, 839.67, 831.57) mm, rotated rx -89.42 ry -19.55 rz -179.75 deg; joints [-74.717, -0.138, 32.721, -170.523, 63.246, -0.126, -170]
  MoveL 983 to (-3457.75, 839.43, 806.57) mm, rotated rx -89.42 ry -19.54 rz -179.74 deg; joints [-74.686, 0.548, 33.096, -169.819, 63.207, -1.375, -170]
  MoveL 984 to (-3457.75, 839.21, 783.57) mm, rotated rx -89.42 ry -19.54 rz -179.74 deg; joints [-74.654, 1.197, 33.425, -169.167, 63.169, -2.528, -170]
  Set speed (1000.0 mm/s)
  MoveL 985 to (-3457.75, 839.21, 783.57) mm, rotated rx -89.42 ry -19.54 rz -179.74 deg; joints [-74.654, 1.197, 33.425, -169.167, 63.169, -2.528, -170]
  MoveL 986 to (-3458.53, 939.2, 782.62) mm, rotated rx -89.42 ry -19.54 rz -179.74 deg; joints [-74.594, -3.237, 37.821, -169.078, 63.082, -2.494, -170]
  Set speed (1000.0 mm/s)
  MoveL 987 to (-3537.75, 940.51, 983.85) mm, rotated rx -89.39 ry -20 rz 179.79 deg; joints [-78.55, -8.488, 34.215, -181.22, 68.827, 8.036, -170]
  MoveL 988 to (-3537.75, 840.51, 984.85) mm, rotated rx -89.39 ry -20 rz 179.79 deg; joints [-78.324, -3.853, 29.992, -180.542, 68.393, 7.568, -170]
  MoveL 989 to (-3537.75, 840.51, 984.85) mm, rotated rx -89.39 ry -20 rz 179.79 deg; joints [-78.324, -3.853, 29.992, -180.542, 68.393, 7.568, -170]
  Set speed (50.0 mm/s)
  MoveL 990 to (-3537.75, 840.56, 990.27) mm, rotated rx -89.39 ry -20 rz 179.79 deg; joints [-78.333, -3.967, 29.883, -180.714, 68.449, 7.823, -170]
  MoveL 991 to (-3537.75, 840.7, 1015.27) mm, rotated rx -89.39 ry -20 rz 179.79 deg; joints [-78.371, -4.475, 29.363, -181.511, 68.718, 8.996, -170]
  MoveL 992 to (-3537.75, 840.82, 1035.38) mm, rotated rx -89.39 ry -21.47 rz 178.33 deg; joints [-77.635, -5.347, 29.092, -179.083, 64.43, 10.312, -170]
  MoveL 993 to (-3537.75, 823.39, 1059.8) mm, rotated rx -125.68 ry 14.5 rz 168.49 deg; joints [-77.516, -4.897, 23.177, -164.712, 68.944, 55.145, -170]
  MoveL 994 to (-3537.75, 805.96, 1084.22) mm, rotated rx -125.72 ry 14.7 rz 168.48 deg; joints [-77.542, -4.416, 21.844, -164.896, 68.836, 56.11, -170]
  MoveL 995 to (-3537.75, 788.53, 1108.64) mm, rotated rx -125.76 ry 14.91 rz 168.47 deg; joints [-77.569, -3.919, 20.499, -165.078, 68.736, 57.074, -170]
  MoveL 996 to (-3537.75, 771.1, 1133.05) mm, rotated rx -125.8 ry 15.13 rz 168.46 deg; joints [-77.596, -3.408, 19.14, -165.256, 68.645, 58.039, -170]
  MoveL 997 to (-3537.75, 753.67, 1157.47) mm, rotated rx -125.85 ry 15.36 rz 168.45 deg; joints [-77.624, -2.881, 17.768, -165.429, 68.561, 59.003, -170]
  MoveL 998 to (-3537.75, 736.24, 1181.89) mm, rotated rx -125.9 ry 15.6 rz 168.43 deg; joints [-77.653, -2.338, 16.383, -165.597, 68.484, 59.967, -170]
  MoveL 999 to (-3537.75, 725.86, 1196.43) mm, rotated rx -125.93 ry 15.75 rz 168.42 deg; joints [-77.67, -2.008, 15.551, -165.693, 68.442, 60.542, -170]
  MoveL 1000 to (-3537.75, 708.33, 1220.78) mm, rotated rx -126.1 ry 16.58 rz 168.37 deg; joints [-77.771, -1.409, 14.216, -165.573, 68.739, 61.468, -170]
  MoveL 1001 to (-3537.75, 690.81, 1245.13) mm, rotated rx -126.29 ry 17.41 rz 168.32 deg; joints [-77.867, -0.798, 12.866, -165.418, 68.996, 62.403, -170]
  MoveL 1002 to (-3537.75, 673.28, 1269.47) mm, rotated rx -126.48 ry 18.24 rz 168.26 deg; joints [-77.957, -0.176, 11.498, -165.228, 69.212, 63.349, -170]
  MoveL 1003 to (-3537.75, 665.41, 1280.4) mm, rotated rx -126.58 ry 18.61 rz 168.23 deg; joints [-77.996, 0.108, 10.879, -165.133, 69.296, 63.778, -170]
  Set speed (1000.0 mm/s)
  MoveL 1004 to (-3537.75, 665.41, 1280.4) mm, rotated rx -126.58 ry 18.61 rz 168.23 deg; joints [-77.996, 0.108, 10.879, -165.133, 69.296, 63.778, -170]
  MoveL 1005 to (-3539.98, 747.91, 1336.88) mm, rotated rx -126.58 ry 18.61 rz 168.23 deg; joints [-78.261, -3.902, 12.71, -166.209, 69.13, 66.254, -170]

--- program second_half_topPaint_startP (robot ABB IRB 5500-27) ---
  Set Ref.: ABB IRB 5500-27 Base
  Set Tool: Paint gun
  MoveJ (second_half_topPaint_app)

--- program first_half_topPaint_startP (robot ABB IRB 5500-27) ---
  Set Ref.: ABB IRB 5500-27 Base
  Set Tool: Paint gun
  MoveJ (first_Half_TopPaint_app)

--- program second_to_First_conn (robot ABB IRB 5500-27) ---
  Set Ref.: ABB IRB 5500-27 Base
  Set Tool: Paint gun
  MoveJ (second_to_home)

--- program CarTopPaintMain (robot ABB IRB 5500-27) ---
  Call second_half_topPaint
  Call second_to_First_conn
  Call first_half_topPaint

--- program sidePaint_startP (robot ABB IRB 5500-27) ---
  Set Ref.: ABB IRB 5500-27 Base
  Set Tool: Paint gun
  MoveJ (sidePaintApp)

--- program CarSidePaintMain (robot ABB IRB 5500-27) ---
  Call side_paint

--- program Home (robot ABB IRB 5500-27) ---
  Set Ref.: ABB IRB 5500-27 Base
  Set Tool: Paint gun
  MoveJ (home)
